Fanuc KAREL source: ke00004.compact.KL

PROGRAM KE00004
%STACKSIZE=65535
%PRIORITY=65535
%NOLOCKGROUP
%ENVIRONMENT REGOPE
VAR
I : INTEGER
S : STRING[80]
STATUS : INTEGER
BEGIN
I=1
S='TEST'
SET_REG_CMT(I,S,STATUS)
END KE00004
